{attribute 'qualified_only'}
{attribute 'strict'}
{attribute 'to_string'}
TYPE E_PolarIIChamberTargetMode :
(
	Disable := 0,
	Manual := 1,
	DryRun := 2,
	Auto := 3
) UINT;
END_TYPE

(* stored: Version 1.1.0.1, ProductVersion 3.1.4026.18
   DUT E_PolarIIChamberTargetMode: Id {14000000-0000-0000-0000-000000000002} *)
